// TIA Portal V21 export
// export: Created 2026-11-10T19:16:33.1871664Z, ExportSetting WithDefaults, DisplayName Totally Integrated Automation Portal, DisplayVersion V21 Update 3, DisplayName STEP 7 Professional, DisplayVersion V21 Update 3, DisplayName STEP 7 Safety, DisplayVersion V21, DisplayName Tech WebApplication, DisplayVersion V21, DisplayName WinCC Basic/Comfort/Advanced, DisplayVersion V21 Update 3, DisplayName WinCC Unified, DisplayVersion V21 Update 3
DATA_BLOCK "FB_300_DB"   // DB2
VERSION : 0.1
// stored: AutoNumber true, InstanceOfName FB_300, InstanceOfType FB
"FB_300"
   // VAR_INPUT
   //    en1 : Bool;
   // END_VAR
   // VAR_OUTPUT
   //    q : Int;
   // END_VAR
   // VAR RETAIN
   //    cnt : Int := 8;
   //    u { S7_SetPoint := 'True'} : "UDT_300";
   // END_VAR
BEGIN
END_DATA_BLOCK
